(* IEC 61131-3 sources: IT-OT/examples, 3 files *)

(* ---- ampel.st ---- *)
(* Fußgängerampel als Schrittkette.
   S7:     Anforderung = DB1.DBX0.0
   OPC UA: ns=2;s=Anforderung *)
PROGRAM Ampel
VAR CONSTANT
  T_GELB  : TIME := T#2s;
  T_ROT   : TIME := T#5s;
  T_RESET : TIME := T#1s;
END_VAR
VAR_INPUT
  Anforderung : BOOL;          (* Taster Fußgänger *)
END_VAR
VAR_OUTPUT
  Auto_Rot, Auto_Gelb, Auto_Gruen : BOOL;
  Fuss_Rot, Fuss_Gruen : BOOL;
  Zyklen : DINT;                (* Anzahl Fußgängerphasen *)
END_VAR
VAR
  Schritt : INT := 0;
  Timer   : TON;
  Taster  : R_TRIG;
  Angefordert : BOOL;
END_VAR

Taster(CLK := Anforderung);
IF Taster.Q THEN
  Angefordert := TRUE;
END_IF;

CASE Schritt OF
  0: (* Autos grün *)
     Auto_Gruen := TRUE; Auto_Gelb := FALSE; Auto_Rot := FALSE;
     Fuss_Rot := TRUE;  Fuss_Gruen := FALSE;
     IF Angefordert THEN
       Schritt := 10;
     END_IF;
  10: (* Autos gelb *)
     Auto_Gruen := FALSE; Auto_Gelb := TRUE;
     Timer(IN := TRUE, PT := T_GELB);
     IF Timer.Q THEN Timer(IN := FALSE); Schritt := 20; END_IF;
  20: (* Autos rot, Fußgänger grün *)
     Auto_Gelb := FALSE; Auto_Rot := TRUE;
     Fuss_Rot := FALSE; Fuss_Gruen := TRUE;
     Timer(IN := TRUE, PT := T_ROT);
     IF Timer.Q THEN Timer(IN := FALSE); Schritt := 30; END_IF;
  30: (* Räumzeit *)
     Fuss_Gruen := FALSE; Fuss_Rot := TRUE;
     Timer(IN := TRUE, PT := T_RESET);
     IF Timer.Q THEN
       Timer(IN := FALSE);
       Angefordert := FALSE;
       Zyklen := Zyklen + 1;
       Schritt := 0;
     END_IF;
ELSE
  Schritt := 0;
END_CASE;
END_PROGRAM

(* ---- foerderband.st ---- *)
(* Förderband mit Teilezählung, Losgröße und Störungsüberwachung. *)
PROGRAM Foerderband
VAR_INPUT
  Start, Stopp, Quittieren : BOOL;
  Sensor_Teil : BOOL;           (* Lichtschranke *)
  Losgroesse  : INT := 10;
END_VAR
VAR_OUTPUT
  Motor   : BOOL;
  Los_Fertig, Stoerung : BOOL;
  Teile   : INT;
  Gesamt  : UDINT;
END_VAR
VAR
  Zaehler : CTU;
  Teil    : R_TRIG;
  Laufzeit_Ohne_Teil : TON;
  Ein     : SR;
END_VAR

Ein(S1 := Start AND NOT Stoerung, R := Stopp OR Stoerung OR Los_Fertig);
Motor := Ein.Q1;

Teil(CLK := Sensor_Teil);
IF Teil.Q THEN Gesamt := Gesamt + 1; END_IF;

Zaehler(CU := Teil.Q, R := Quittieren, PV := Losgroesse);
Teile := Zaehler.CV;
Los_Fertig := Zaehler.Q;

(* Störung: Band läuft 10 s ohne dass ein Teil erkannt wird *)
Laufzeit_Ohne_Teil(IN := Motor AND NOT Sensor_Teil, PT := T#10s);
IF Laufzeit_Ohne_Teil.Q THEN
  Stoerung := TRUE;
END_IF;
IF Quittieren THEN
  Stoerung := FALSE;
END_IF;
END_PROGRAM

(* ---- tank.st ---- *)
(* Füllstandsregelung mit Zweipunktregler und simulierter Strecke.
   Ideal zum Testen von HMI/SCADA-Anbindungen über S7 oder OPC UA. *)
PROGRAM Tank
VAR_INPUT
  Automatik : BOOL := TRUE;
  Sollwert  : REAL := 60.0;    (* % *)
  Hysterese : REAL := 5.0;     (* % *)
  Abfluss   : REAL := 0.15;    (* %/Zyklus *)
END_VAR
VAR_OUTPUT
  Fuellstand : REAL := 20.0;   (* % *)
  Pumpe      : BOOL;
  Alarm_Hoch, Alarm_Tief : BOOL;
  Pumpenstarts : DINT;
END_VAR
VAR
  Zufluss : REAL := 0.4;
  Start   : R_TRIG;
  Alarm_Verz : TON;
END_VAR

IF Automatik THEN
  IF Fuellstand < Sollwert - Hysterese THEN
    Pumpe := TRUE;
  ELSIF Fuellstand > Sollwert + Hysterese THEN
    Pumpe := FALSE;
  END_IF;
END_IF;

Start(CLK := Pumpe);
IF Start.Q THEN Pumpenstarts := Pumpenstarts + 1; END_IF;

(* Simulation der Strecke *)
IF Pumpe THEN
  Fuellstand := Fuellstand + Zufluss;
END_IF;
Fuellstand := LIMIT(0.0, Fuellstand - Abfluss, 100.0);

Alarm_Verz(IN := Fuellstand > 95.0 OR Fuellstand < 5.0, PT := T#2s);
Alarm_Hoch := Alarm_Verz.Q AND Fuellstand > 95.0;
Alarm_Tief := Alarm_Verz.Q AND Fuellstand < 5.0;
END_PROGRAM
